FUNCTION_BLOCK FB_DomeControl IMPLEMENTS I_Dome
VAR_INPUT
	ipTelescope: I_RaDecTelescope;
END_VAR
VAR
	ipState		: I_DomeState := fbDomeIdleState;
	bOpen		: BOOL;
	bClose		: BOOL;
	bReset		: BOOL;
	bHome		: BOOL;
	bTrack		: BOOL;
	bPark		: BOOL;
	bStop		: BOOL;
	bStopDone	: BOOL;
	
	fDomeAziGoInput			: LREAL := 180.0;
	fDomeAziGo				: LREAL := 180.0;
	fDomeAziCurrent			: LREAL := 0.0;
	eDomeRotationState		: E_DomeRotationState;
	eDomeRotationStateOld	: E_DomeRotationState;
	eDomeShutterState		: E_RoofState;
	eDomeShutterStateOld	: E_RoofState;
	bParked			: BOOL;
	
	bDomeError	: BOOL;
	iDomeErrorID: UINT;
	
	ipStateOld			: I_DomeState := fbDomeIdleState;
	fbDomeCloseingState : FB_DomeClosingState(THIS);
	fbDomeErrorState	: FB_DomeErrorState(THIS);
	fbDomeHomeingState	: FB_DomeHomingState(THIS);
	fbDomeIdleState		: FB_DomeIdleState(THIS);
	fbDomeOpeningState	: FB_DomeOpeningState(THIS);
	fbDomeMovingState	: FB_DomeMovingState(THIS);
	fbDomeParkingState	: FB_DomeParkingState(THIS);
	fbDomeStoppingState	: FB_DomeStoppingState(THIS);
	

	rtrigOpen		: R_TRIG;
	rtrigClose		: R_TRIG;
	rtrigReset		: R_TRIG;
	rtrigHome		: R_TRIG;
	rtrigPark		: R_TRIG;
	rtrigStop		: R_TRIG;
	
	fbComm			: I_Comm;
	tonComm 		: TON := (PT:=T#5S);
	
	fbDomeParkedEvent:	FB_EventLog;
	fbDomeStopEvent:	FB_EventLog;
	fbDomeErrorEvent: FB_EventLog;
	
	sSendstring	: STRING;
	Stage		: UINT:= 0;
	Timer		: TON := (PT:=T#30S);
	fbSend		: SendString;
	bSendBusy	: BOOL;
	eSendErrorID: ComError_t;

	fbReceive		: ReceiveString;
	sReceivedString	: STRING;
	sLastReceivedString: STRING;
	bStringReceived	: BOOL;
	bReceiveBusy	: BOOL;
	bReceiveError	: BOOL;
	eReceiveErrorID	: ComError_t;
	bReceiveTimeout	: BOOL;
END_VAR
VAR CONSTANT
	nCapabilities : INT := 2; 	//OPEN TSI : TELESCOPE.CONFIG.CAPABILITIES
END_VAR

// account for off center mount
IF fDomeAziGoInput >= 0.0 AND fDomeAziGoInput < 115.0 THEN
	fDomeAziGo := fDomeAziGoInput - 5.0;
ELSIF fDomeAziGoInput >= 225.0 AND fDomeAziGoInput < 360.0 THEN
	fDomeAziGo := fDomeAziGoInput + 5.0;
ELSE
	fDomeAziGo := fDomeAziGoInput;
END_IF

//	Receive string data:
fbReceive(
	Prefix:='',
	Suffix:= '',
	Timeout:= T#1S,
	ReceivedString:= sReceivedString,
	RXbuffer:= RxBufferDome,
	StringReceived=> bStringReceived,
	Busy=> bReceiveBusy,
	Error=> ,
	RxTimeout=> bReceiveTimeout );
// Check Errors
IF fbSend.Error <> COMERROR_NOERROR THEN
	eSendErrorID := fbSend.Error;
	bDomeError := TRUE;
END_IF
IF fbReceive.Error <> COMERROR_NOERROR THEN
	eReceiveErrorID := fbReceive.Error;
	bDomeError := TRUE;
END_IF

IF bDomeError THEN
	THIS^.ipState.FoundError();
END_IF

rtrigOpen(CLK := bOpen);
rtrigClose(CLK := bClose);
rtrigReset(CLK := bReset);
rtrigHome(CLK := bHome);
rtrigPark(CLK := bPark);
rtrigStop(CLK := bStop);

// #96: a stop wins over every other request of the same scan, which are dropped with it
IF (rtrigStop.Q) THEN
	bStop := FALSE;
	bOpen := FALSE;
	bClose := FALSE;
	bHome := FALSE;
	bPark := FALSE;
	bTrack := FALSE;
	ipState.StopCommand();
END_IF

IF (rtrigReset.Q) THEN
	bReset := FALSE;
	ipState.ResetCommand();
END_IF

IF (rtrigClose.Q) THEN
	bClose := FALSE;
	ipState.CloseCommand();
END_IF

IF (rtrigOpen.Q) THEN
	bOpen := FALSE;
	ipState.OpenCommand();
END_IF

IF (rtrigHome.Q) THEN
	bHome := FALSE;
	ipState.HomeCommand();
END_IF

IF (rtrigPark.Q) THEN
	bPark := FALSE;
	bTrack := FALSE;
	ipState.ParkCommand();
END_IF

// #83: requests are one-shot, like the covers (#66). They are consumed in this scan whether they produced an edge or
// not: a caller repeating a request every scan gave a single edge and then left the flag TRUE, so no later request of
// that kind had an edge until a PLC restart.
bOpen := FALSE;
bClose := FALSE;
bReset := FALSE;
bHome := FALSE;
bPark := FALSE;
bStop := FALSE;

bStopDone := FALSE;
ipState.RunState();

IF eDomeRotationState = E_DomeRotationState.parked AND eDomeShutterState = E_RoofState.closed THEN
	bParked := TRUE;
ELSE
	bParked := FALSE;
END_IF
// send telemetry
tonComm(IN:=TRUE);
IF tonComm.Q THEN // publish new payload every 5 seconds
	tonComm(IN:=FALSE);
	THIS^._SendTelemetry();	
END_IF


fbDomeParkedEvent(
	Trigger := bParked,
	Level := ADSLOG_MSGTYPE_HINT,
	OnMessage := 'Dome is in parking position and closed.',
	comm:= fbComm);
fbDomeStopEvent(
	Trigger := bStopDone,
	Level := ADSLOG_MSGTYPE_HINT,
	OnMessage := 'Dome stopped: rotation holds the current azimuth, a shutter movement is not stopped.',
	comm:= fbComm);
fbDomeErrorEvent(
	Trigger := bDomeError,
	Level := ADSLOG_MSGTYPE_ERROR,
	FormatString := 'Dome Error %s',
	OnMessage := 'found.',
	OffMessage := 'resolved.',
	comm:= fbComm);
// Buffer
ipStateOld := ipState;
eDomeRotationStateOld := eDomeRotationState;
eDomeShutterStateOld := eDomeShutterState;

PROPERTY _DomeRotationState : E_DomeRotationState
GET
_DomeRotationState := eDomeRotationState;
END_GET
SET
eDomeRotationState := _DomeRotationState;
END_SET
END_PROPERTY

PROPERTY _DomeShutterState : E_RoofState
GET
_DomeShutterState := eDomeShutterState;
END_GET
SET
eDomeShutterState := _DomeShutterState;
END_SET
END_PROPERTY

PROPERTY  _Error : BOOL
GET
_Error := bDomeError;
END_GET
SET
bDomeError := _Error;
END_SET
END_PROPERTY

PROPERTY _StopDone : BOOL
GET
_StopDone := bStopDone;
END_GET
SET
bStopDone := _StopDone;
END_SET
END_PROPERTY

PROPERTY _HasReceivedString : Bool
GET
_HasReceivedString := bStringReceived;
END_GET
SET
END_SET
END_PROPERTY

PROPERTY _Parked : BOOL
GET
_Parked := bParked;
END_GET
SET
bParked := _Parked;
END_SET
END_PROPERTY

PROPERTY _Position : LREAL
GET
_Position := fDomeAziGo;
END_GET
SET
fDomeAziCurrent := _Position;
END_SET
END_PROPERTY

PROPERTY _ReceivedString : STRING
GET
_ReceivedString := sReceivedString;
END_GET
SET
END_SET
END_PROPERTY

METHOD _SendTelemetry : BOOL
VAR_INPUT
END_VAR
IF eDomeShutterState = E_RoofState.opened THEN
	fbComm.PublishLREAL('telescope', 'dome', 'AUXILIARY.DOME.REALPOS', 1.0);
ELSIF eDomeShutterState = E_RoofState.closing OR eDomeShutterState = E_RoofState.opening OR eDomeShutterState = E_RoofState.unknown THEN
	fbComm.PublishLREAL('telescope', 'dome', 'AUXILIARY.DOME.REALPOS', 0.5);
ELSIF eDomeShutterState = E_RoofState.closed THEN
	fbComm.PublishLREAL('telescope', 'dome', 'AUXILIARY.DOME.REALPOS', 0.0);
ELSE
	fbComm.PublishLREAL('telescope', 'dome', 'AUXILIARY.DOME.REALPOS', -1.0);
END_IF

IF ipState.StateID = 'Opening State' THEN
	fbComm.PublishLREAL('telescope', 'dome', 'AUXILIARY.DOME.TARGETPOS', 1.0);
ELSE
	fbComm.PublishLREAL('telescope', 'dome', 'AUXILIARY.DOME.TARGETPOS', 0.0);
END_IF

IF bDomeError THEN
	fbComm.PublishINT('telescope', 'dome', 'AUXILIARY.DOME.ERROR_STATE', 1);
	fbComm.PublishLREAL('telescope', 'dome', 'AUXILIARY.DOME.READY_STATE', -1.0);
ELSE
	fbComm.PublishINT('telescope', 'dome', 'AUXILIARY.DOME.ERROR_STATE', 0);
	IF bParked THEN
		fbComm.PublishLREAL('telescope', 'dome', 'AUXILIARY.DOME.READY_STATE', 0.0);
	ELSIF bTrack THEN
		fbComm.PublishLREAL('telescope', 'dome', 'AUXILIARY.DOME.READY_STATE', 8.0);
	ELSE
		fbComm.PublishLREAL('telescope', 'dome', 'AUXILIARY.DOME.READY_STATE', 1.0);
	END_IF
END_IF

IF eDomeRotationState = E_DomeRotationState.slewing OR eDomeRotationState = E_DomeRotationState.unknown THEN
	fbComm.PublishLREAL('telescope', 'dome', 'AUXILIARY.DOME.MOTION_STATE', 1.0);
ELSE
	fbComm.PublishLREAL('telescope', 'dome', 'AUXILIARY.DOME.MOTION_STATE', 0.0);
END_IF
fbComm.PublishLREAL('telescope', 'dome', 'AUXILIARY.DOME.AZ', THIS^.Position);
END_METHOD

PROPERTY _Track : BOOL
GET
_Track := bTrack;
END_GET
END_PROPERTY

PROPERTY Capabilities : INT
GET
Capabilities := nCapabilities;
END_GET
END_PROPERTY

METHOD Close : BOOL
VAR_INPUT
END_VAR
bClose:=True;
END_METHOD

PROPERTY Closed : BOOL
GET
END_GET
END_PROPERTY

PROPERTY Error : Bool
GET
Error := bDomeError;
END_GET
END_PROPERTY

PROPERTY ErrorID : UDINT
GET
END_GET
END_PROPERTY

//FB_Init is always available implicitly and it is used primarily for initialization.
//The return value is not evaluated. For a specific influence, you can also declare the
//methods explicitly and provide additional code there with the standard initialization
//code. You can evaluate the return value.
METHOD FB_Init: BOOL
VAR_INPUT
    bInitRetains	: BOOL; // TRUE: the retain variables are initialized (reset warm / reset cold)
    bInCopyCode		: BOOL;  // TRUE: the instance will be copied to the copy code afterward (online change)
	comm			: I_Comm;
END_VAR
THIS^.fbComm 				:= comm;
END_METHOD

METHOD Open : BOOL
VAR_INPUT
END_VAR
bOpen := True;
END_METHOD

PROPERTY Opened : BOOL
GET
END_GET
END_PROPERTY

METHOD Park : BOOL
VAR_INPUT
END_VAR
bPark := TRUE;
END_METHOD

PROPERTY Parked : BOOL
GET
Parked := bParked;
END_GET
END_PROPERTY

PROPERTY Position : LREAL
GET
Position := fDomeAziCurrent;
END_GET
SET
fDomeAziGoInput := Position;
END_SET
END_PROPERTY

METHOD Reset : BOOL
VAR_INPUT
END_VAR
bReset := True;
END_METHOD

PROPERTY RotState : E_DomeRotationState
GET
RotState := eDomeRotationState;
END_GET
END_PROPERTY

METHOD SetState : BOOL
VAR_INPUT
	newState :I_DomeState;
END_VAR
THIS^.ipState := newState;
END_METHOD

{warning 'add property implementation'}
PROPERTY ShutterState : BROTLib.E_RoofState
GET
END_GET
SET
END_SET
END_PROPERTY

PROPERTY Slewing : BOOL
GET
END_GET
END_PROPERTY

METHOD Stop : BOOL
VAR_INPUT
END_VAR
// #96: the dome has no stop command, the state holds the azimuth it reads (FB_DomeStoppingState)
bStop := TRUE;
END_METHOD

METHOD StopTrack : BOOL
VAR_INPUT
END_VAR
bTrack := FALSE;
END_METHOD

METHOD Track : BOOL
VAR_INPUT
END_VAR
bTrack := TRUE;
END_METHOD

PROPERTY Tracking : BOOL
GET
Tracking := bTrack;
END_GET
END_PROPERTY

END_FUNCTION_BLOCK

(* stored: Version 1.1.0.1, ProductVersion 3.1.4024.15
   POU FB_DomeControl: Id {6d19e4e0-cd8e-40f8-8605-b776152ffcc0}, SpecialFunc None
   Folder internal properties: Id {f2b50677-3a48-4dff-8e4d-06640225c481}
   Folder properties: Id {aebe3fd9-357f-41e3-8c30-105b311d4951}
   Property _DomeRotationState: Id {94e281da-2d55-4137-b423-8bf7bc330143}
   Get Get: Id {e931b510-c0b8-460e-90fe-ec0def1d87ff}
   Set Set: Id {444b45a3-ce96-43fc-b5d3-4fd60b06192b}
   Property _DomeShutterState: Id {5d37da6d-da48-4528-837f-be475da99739}
   Get Get: Id {3e09792f-5402-466e-8155-6362efadc1a5}
   Set Set: Id {b69684dc-6640-4585-a298-28b78eac4adb}
   Property _Error: Id {c93dc26f-1216-4281-a3a2-0ba8e3029faf}
   Get Get: Id {766ee077-f5ca-4c10-8364-d6db87eb6439}
   Set Set: Id {e7ecb5f9-adba-48a7-aafb-40be532480f0}
   Property _StopDone: Id {972f1c99-75d8-4fff-ae5d-301663a13d0f}
   Get Get: Id {e95f46bc-fd74-4b65-8b40-76498780211b}
   Set Set: Id {f7672a6c-da04-4be5-bce4-44adb61d318d}
   Property _HasReceivedString: Id {efe4ec58-b013-4bd3-91d7-a40e68ac61d6}
   Get Get: Id {6af32aed-d4e7-435f-a147-9af66e31cbf3}
   Set Set: Id {82b0d852-aa2b-4f8d-8a49-7fbd2bfaec1c}
   Property _Parked: Id {1b15552c-bfee-42da-88e4-7dcb176a1825}
   Get Get: Id {ce33e28b-4dd6-4d2b-bf76-aba9b91ad629}
   Set Set: Id {4c46eccf-1f31-4481-83e7-6180d7889bee}
   Property _Position: Id {ae105779-0aa0-4d2f-821e-0f47310d89e1}
   Get Get: Id {0c9924d3-2af6-4b94-83fc-e627953dfa21}
   Set Set: Id {651597fa-a85f-49cd-8330-7278a65501fd}
   Property _ReceivedString: Id {ff9987e3-3e05-4fae-a5e0-cb86b6b8209d}
   Get Get: Id {caa6b28d-538c-43d7-8264-8d51b155f525}
   Set Set: Id {d34cb6a8-9699-4b13-9e1d-7c89f67e2095}
   Method _SendTelemetry: Id {fbbd6c37-f392-4c14-80af-cf2ffd3d50c5}
   Property _Track: Id {a690fc2a-3ca4-499b-bcfe-9a72b5ec9057}
   Get Get: Id {64355058-626f-404d-8e97-1c1fd171de1e}
   Property Capabilities: Id {a5232eb4-5866-434a-858f-b0136e7dd593}
   Get Get: Id {97d77058-b27e-4c1e-ab84-3307e1bea0b7}
   Method Close: Id {df2077f2-da90-4613-b060-6d6c3ae4fa51}
   Property Closed: Id {6d997260-0381-44c8-9f75-ce63c1cb4011}
   Get Get: Id {748e5a80-31e8-4286-bfa0-1a642c517ee7}
   Property Error: Id {268476f6-d236-45b6-8bd2-428f6ed1c5c5}
   Get Get: Id {1e94d00a-28b4-4617-af13-fff028d77e00}
   Property ErrorID: Id {e66424b4-fdaf-4b3d-92ec-390d6ab9acbb}
   Get Get: Id {1eb8ee0b-47e9-4214-bdd5-d2740de92e5f}
   Method FB_Init: Id {0ad2fe54-2f8b-455c-ac43-fce68b95c2e8}
   Method Open: Id {06a72384-aba2-42e8-9b34-7edb45f49723}
   Property Opened: Id {65547067-38a4-4670-ad36-0884355dc8d3}
   Get Get: Id {f8408426-5aa1-4ac5-8fa2-912147109708}
   Method Park: Id {3be05401-3914-4f1f-9af7-03ba8643ddec}
   Property Parked: Id {e400500f-7f31-4456-b38c-60e2d41191a1}
   Get Get: Id {b243146e-6556-4e7d-843a-c7cbc2974276}
   Property Position: Id {566a0c40-7cf6-4687-b475-98742f4a3e93}
   Get Get: Id {51596a5f-29ff-4600-84cd-814b0fa48e76}
   Set Set: Id {ac1cf9b5-c5c0-487f-baa8-762c0c8e8d55}
   Method Reset: Id {64e6a766-3201-41a9-a8b3-86ae4ee59491}
   Property RotState: Id {8c2c601e-a673-493f-a0e6-8cb4c126be63}
   Get Get: Id {1b5f019c-56a3-4acd-86fa-be8fed03a696}
   Method SetState: Id {bac7998a-96e0-484d-9b0b-984b4f2ae380}
   Property ShutterState: Id {5fd910c8-e41a-4706-b0a5-896ca2b3fba0}
   Get Get: Id {cd0a457a-ce60-4149-bafe-b923afc36585}
   Set Set: Id {366d60c6-d226-4cf0-928a-a262b9375329}
   Property Slewing: Id {f4557448-d077-4c28-8ed8-f77cf26bab9c}
   Get Get: Id {b28436fa-18d0-4eee-9d60-f0af07e234ec}
   Method Stop: Id {437563e5-1f1f-4c46-b138-d206b8d0b2ae}
   Method StopTrack: Id {592d7f7e-1fdb-4ea9-b619-2542fb2b964e}
   Method Track: Id {098e5b71-cc16-4ffe-ab71-96c1984155a2}
   Property Tracking: Id {1a2cedbc-ec50-4d4c-88f2-62da93b16706}
   Get Get: Id {6f0c9f90-dee6-4c1b-b31b-03a846e8a5b2} *)
